(* Logix 5000 project; controller TFF vendor 1 type 14 code 107 rev 34.11; software revision 34.03; part 19 of 36 *)
(* tags used below, declared in another part *)
   AddressPump1 : DINT;   // Temp Address for Pump 1
   AddressPump2 : DINT;   // Temp Address for Pump 2
   Index : DINT;   // Index
   AlarmAnalog : AlarmAnalog[50];   // Analog Alarm Array
   AlarmControl : AlarmControl;   // Alarm Control
   AlarmDeviation : AlarmDeviation[20];   // Control Loop Deviation Alarm Array
   AnalogPoint : AnalogInput[50];   // Analog Input Array
   ControlLoop : ControlLoop[20];   // Control Loop Array
   ControlLoop_FeedBagLevel : ALIAS FOR ControlLoop[2];   // Feed Bag Level Control Loop
   ControlLoop_FeedBagLevelAlarm : ALIAS FOR AlarmDeviation[2];   // Feed Bag Level Control Loop Deviation Alarm
   ControlLoop_FeedPump : ALIAS FOR ControlLoop[1];   // Feed Pump Control Loop
   ControlLoop_FeedPumpAlarm : ALIAS FOR AlarmDeviation[1];   // Feed Pump Control Loop Deviation Alarm
   ControlLoop_PCV001 : ALIAS FOR ControlLoop[3];   // PCV001 Control Loop
   ControlLoop_PCV001Alarm : ALIAS FOR AlarmDeviation[3];   // PCV001 Control Loop Deviation Alarm
   ControlLoop_PCV101 : ALIAS FOR ControlLoop[5];   // PCV101 Control Loop
   ControlLoop_PCV101Alarm : ALIAS FOR AlarmDeviation[5];   // PCV101 Control Loop Deviation Alarm
   Drive : Drive[11];   // Drives Array
   PCV001 : ALIAS FOR AnalogPoint[3];   // Retentate Pressure Control Valve Position
   PCV101 : ALIAS FOR AnalogPoint[4];   // Filtrate Pressure Control Valve Position
   Timers : Timers[22];   // Timer Array
(* Process, continued *)

ROUTINE Alarm_Analog   (* ladder *)
// Analog Alarm Routine
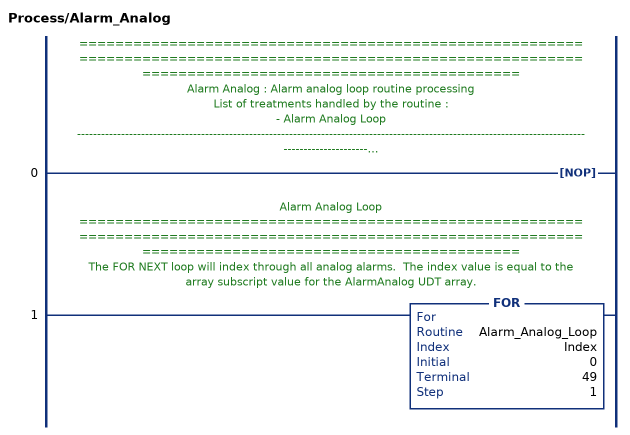
   // ==========================================================================================================================================================
   //                                                                                                                 Alarm Analog : Alarm analog loop routine processing
   //                                                     List of treatments handled by the routine :
   //                                                          - Alarm Analog Loop
   //                                                     -----------------------------------------------------------------------------------------------------------------------------------------------------
   //                                                     History
   //                                                          2019-AUG-13 - Actemium - B. Roch - Initial version for Candidate Release 3.00.00.00.a
   // ==========================================================================================================================================================
   0: NOP();
   // Alarm Analog Loop
   // ==========================================================================================================================================================
   // The FOR NEXT loop will index through all analog alarms.  The index value is equal to the array subscript value for the AlarmAnalog UDT array.
   1: FOR(Alarm_Analog_Loop,Index,0,49,1);
END_ROUTINE

ROUTINE Alarm_Analog_Loop   (* ladder *)
// Analog Alarm Routine
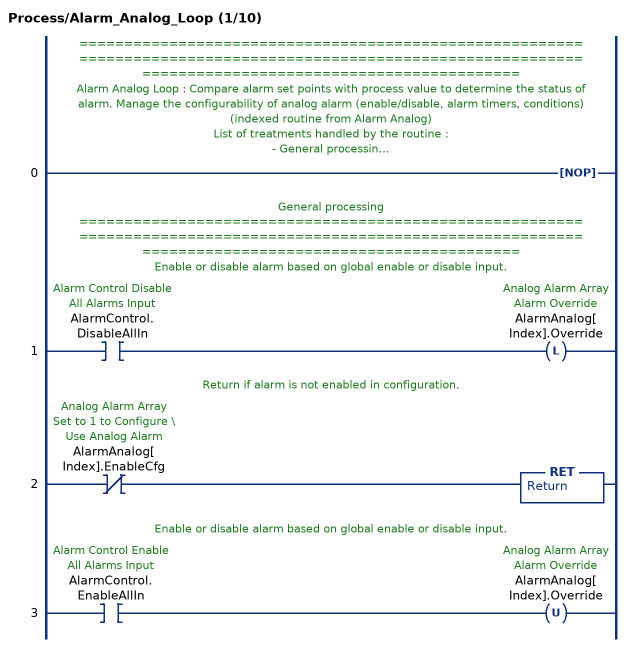
   // ==========================================================================================================================================================
   //           Alarm Analog Loop : Compare alarm set points with process value to determine the status of alarm. Manage the configurability of analog alarm (enable/disable, alarm timers, conditions)
   //                                                                                                                             (indexed routine from Alarm Analog)
   //                                                     List of treatments handled by the routine :
   //                                                          - General processing
   //                                                          - Alarm Acknowledged status
   //                                                          - Alarm conditioned on pump operating status
   //                                                          - Alarm LOLO processing
   //                                                          - Alarm LO processing
   //                                                          - Alarm HI processing
   //                                                          - Alarm HIHI processing
   //                                                          - Alarm status processing
   //                                                     -----------------------------------------------------------------------------------------------------------------------------------------------------
   //                                                     History
   //                                                          2019-AUG-13 - Actemium - B. Roch - Initial version for Candidate Release 3.00.00.00.a
   // ==========================================================================================================================================================
   0: NOP();
   // General processing
   // ==========================================================================================================================================================
   // Enable or disable alarm based on global enable or disable input.
   1: XIC(AlarmControl.DisableAllIn)OTL(AlarmAnalog[Index].Override);
   // Return if alarm is not enabled in configuration.
   2: XIO(AlarmAnalog[Index].EnableCfg)RET();
   // Enable or disable alarm based on global enable or disable input.
   3: XIC(AlarmControl.EnableAllIn)OTU(AlarmAnalog[Index].Override);
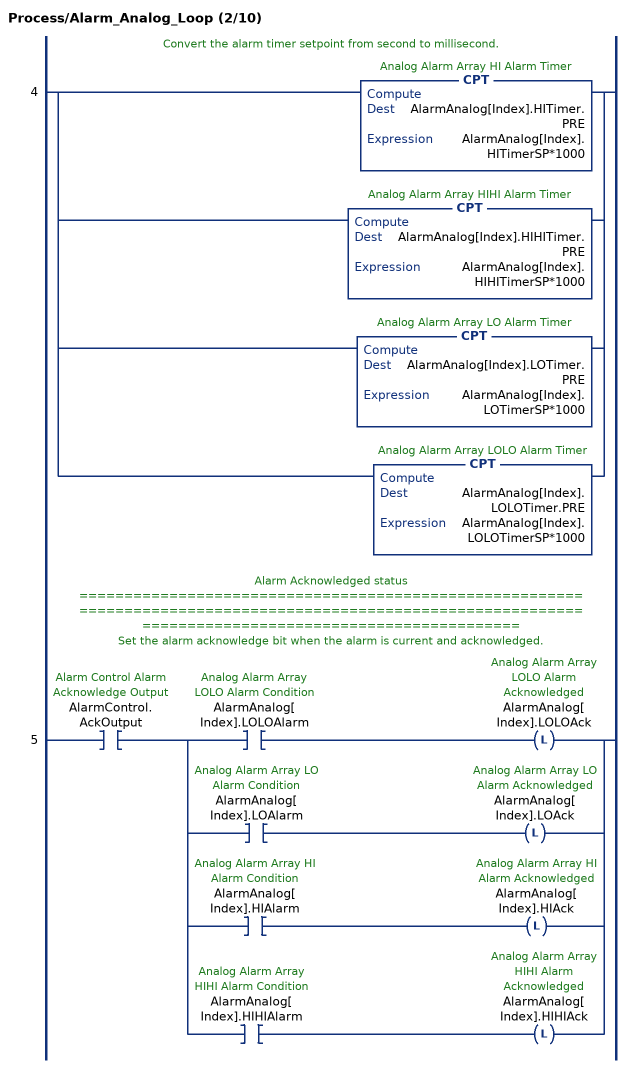
   // Convert the alarm timer setpoint from second to millisecond.
   4: [CPT(AlarmAnalog[Index].HITimer.PRE,AlarmAnalog[Index].HITimerSP*1000) ,CPT(AlarmAnalog[Index].HIHITimer.PRE,AlarmAnalog[Index].HIHITimerSP*1000) ,CPT(AlarmAnalog[Index].LOTimer.PRE,AlarmAnalog[Index].LOTimerSP*1000) ,CPT(AlarmAnalog[Index].LOLOTimer.PRE,AlarmAnalog[Index].LOLOTimerSP*1000) ];
   // Alarm Acknowledged status
   // ==========================================================================================================================================================
   // Set the alarm acknowledge bit when the alarm is current and acknowledged.
   5: XIC(AlarmControl.AckOutput)[XIC(AlarmAnalog[Index].LOLOAlarm) OTL(AlarmAnalog[Index].LOLOAck) ,XIC(AlarmAnalog[Index].LOAlarm) OTL(AlarmAnalog[Index].LOAck) ,XIC(AlarmAnalog[Index].HIAlarm) OTL(AlarmAnalog[Index].HIAck) ,XIC(AlarmAnalog[Index].HIHIAlarm) OTL(AlarmAnalog[Index].HIHIAck) ];
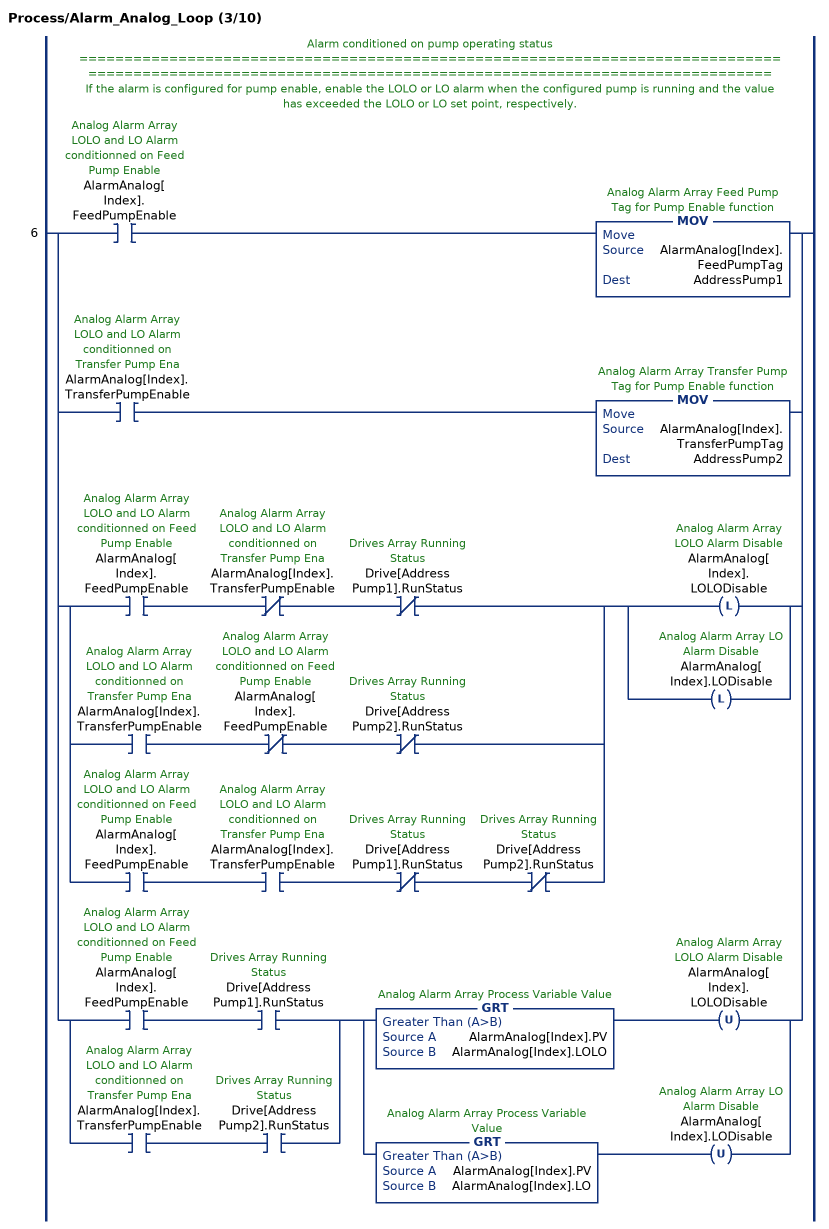
   // Alarm conditioned on pump operating status
   // ==========================================================================================================================================================
   // If the alarm is configured for pump enable, enable the LOLO or LO alarm when the configured pump is running and the value has exceeded the LOLO or LO set point, respectively.
   6: [XIC(AlarmAnalog[Index].FeedPumpEnable) MOV(AlarmAnalog[Index].FeedPumpTag,AddressPump1) ,XIC(AlarmAnalog[Index].TransferPumpEnable) MOV(AlarmAnalog[Index].TransferPumpTag,AddressPump2) ,[XIC(AlarmAnalog[Index].FeedPumpEnable) XIO(AlarmAnalog[Index].TransferPumpEnable) XIO(Drive[AddressPump1].RunStatus) ,XIC(AlarmAnalog[Index].TransferPumpEnable) XIO(AlarmAnalog[Index].FeedPumpEnable) XIO(Drive[AddressPump2].RunStatus) ,XIC(AlarmAnalog[Index].FeedPumpEnable) XIC(AlarmAnalog[Index].TransferPumpEnable) XIO(Drive[AddressPump1].RunStatus) XIO(Drive[AddressPump2].RunStatus) ] [OTL(AlarmAnalog[Index].LOLODisable) ,OTL(AlarmAnalog[Index].LODisable) ] ,[XIC(AlarmAnalog[Index].FeedPumpEnable) XIC(Drive[AddressPump1].RunStatus) ,XIC(AlarmAnalog[Index].TransferPumpEnable) XIC(Drive[AddressPump2].RunStatus) ] [GRT(AlarmAnalog[Index].PV,AlarmAnalog[Index].LOLO) OTU(AlarmAnalog[Index].LOLODisable) ,GRT(AlarmAnalog[Index].PV,AlarmAnalog[Index].LO) OTU(AlarmAnalog[Index].LODisable) ] ];
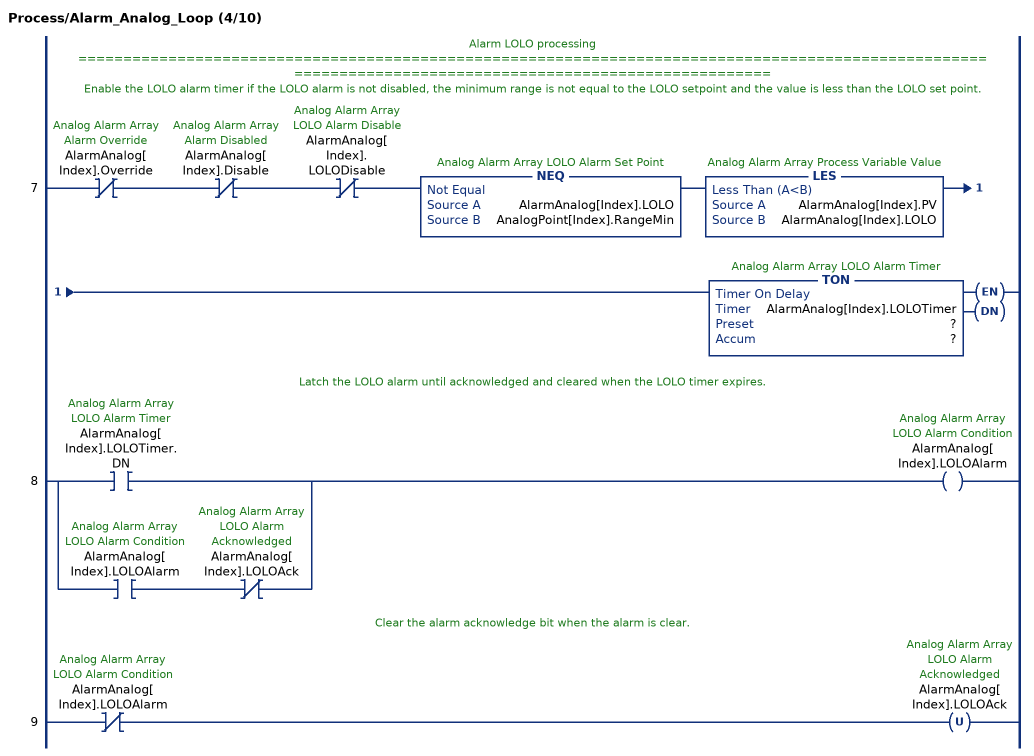
   // Alarm LOLO processing
   // ==========================================================================================================================================================
   // Enable the LOLO alarm timer if the LOLO alarm is not disabled, the minimum range is not equal to the LOLO setpoint and the value is less than the LOLO set point.
   7: XIO(AlarmAnalog[Index].Override)XIO(AlarmAnalog[Index].Disable)XIO(AlarmAnalog[Index].LOLODisable)NEQ(AlarmAnalog[Index].LOLO,AnalogPoint[Index].RangeMin)LES(AlarmAnalog[Index].PV,AlarmAnalog[Index].LOLO)TON(AlarmAnalog[Index].LOLOTimer,?,?);
   // Latch the LOLO alarm until acknowledged and cleared when the LOLO timer expires.
   8: [XIC(AlarmAnalog[Index].LOLOTimer.DN) ,XIC(AlarmAnalog[Index].LOLOAlarm) XIO(AlarmAnalog[Index].LOLOAck) ]OTE(AlarmAnalog[Index].LOLOAlarm);
   // Clear the alarm acknowledge bit when the alarm is clear.
   9: XIO(AlarmAnalog[Index].LOLOAlarm)OTU(AlarmAnalog[Index].LOLOAck);
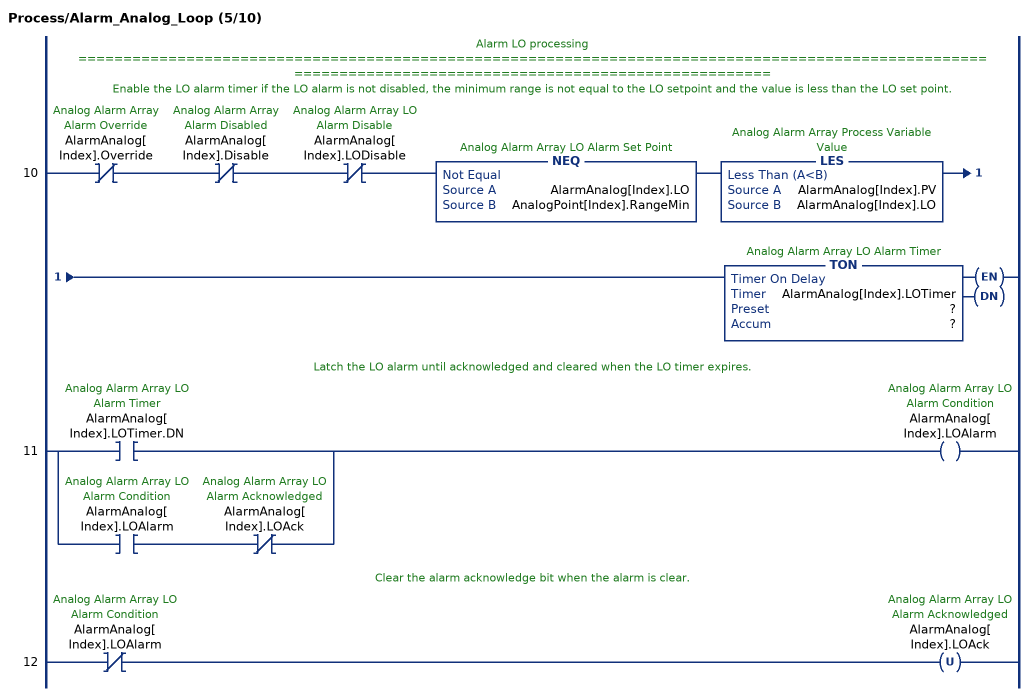
   // Alarm LO processing
   // ==========================================================================================================================================================
   // Enable the LO alarm timer if the LO alarm is not disabled, the minimum range is not equal to the LO setpoint and the value is less than the LO set point.
   10: XIO(AlarmAnalog[Index].Override)XIO(AlarmAnalog[Index].Disable)XIO(AlarmAnalog[Index].LODisable)NEQ(AlarmAnalog[Index].LO,AnalogPoint[Index].RangeMin)LES(AlarmAnalog[Index].PV,AlarmAnalog[Index].LO)TON(AlarmAnalog[Index].LOTimer,?,?);
   // Latch the LO alarm until acknowledged and cleared when the LO timer expires.
   11: [XIC(AlarmAnalog[Index].LOTimer.DN) ,XIC(AlarmAnalog[Index].LOAlarm) XIO(AlarmAnalog[Index].LOAck) ]OTE(AlarmAnalog[Index].LOAlarm);
   // Clear the alarm acknowledge bit when the alarm is clear.
   12: XIO(AlarmAnalog[Index].LOAlarm)OTU(AlarmAnalog[Index].LOAck);
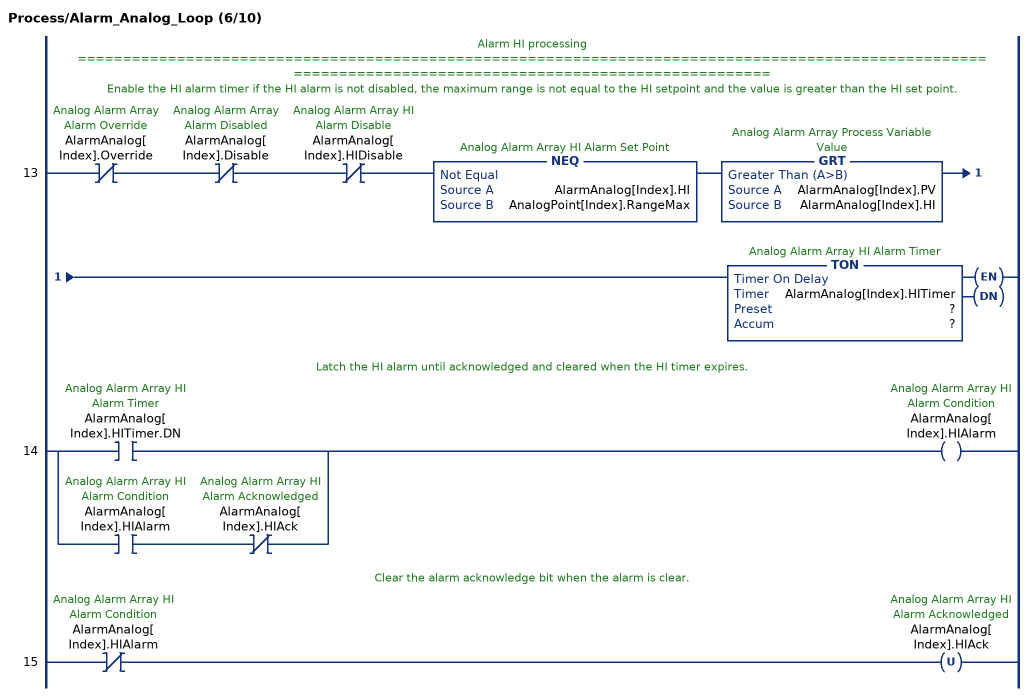
   // Alarm HI processing
   // ==========================================================================================================================================================
   // Enable the HI alarm timer if the HI alarm is not disabled, the maximum range is not equal to the HI setpoint and the value is greater than the HI set point.
   13: XIO(AlarmAnalog[Index].Override)XIO(AlarmAnalog[Index].Disable)XIO(AlarmAnalog[Index].HIDisable)NEQ(AlarmAnalog[Index].HI,AnalogPoint[Index].RangeMax)GRT(AlarmAnalog[Index].PV,AlarmAnalog[Index].HI)TON(AlarmAnalog[Index].HITimer,?,?);
   // Latch the HI alarm until acknowledged and cleared when the HI timer expires.
   14: [XIC(AlarmAnalog[Index].HITimer.DN) ,XIC(AlarmAnalog[Index].HIAlarm) XIO(AlarmAnalog[Index].HIAck) ]OTE(AlarmAnalog[Index].HIAlarm);
   // Clear the alarm acknowledge bit when the alarm is clear.
   15: XIO(AlarmAnalog[Index].HIAlarm)OTU(AlarmAnalog[Index].HIAck);
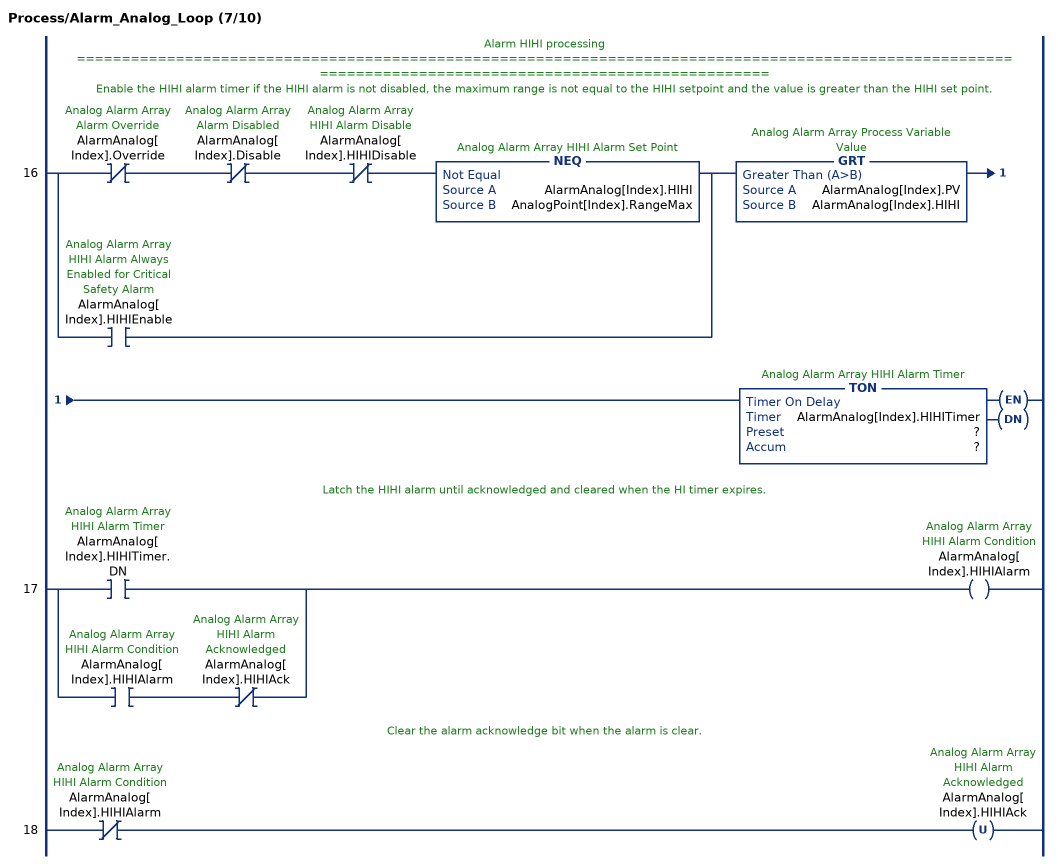
   // Alarm HIHI processing
   // ==========================================================================================================================================================
   // Enable the HIHI alarm timer if the HIHI alarm is not disabled, the maximum range is not equal to the HIHI setpoint and the value is greater than the HIHI set point.
   16: [XIO(AlarmAnalog[Index].Override) XIO(AlarmAnalog[Index].Disable) XIO(AlarmAnalog[Index].HIHIDisable) NEQ(AlarmAnalog[Index].HIHI,AnalogPoint[Index].RangeMax) ,XIC(AlarmAnalog[Index].HIHIEnable) ]GRT(AlarmAnalog[Index].PV,AlarmAnalog[Index].HIHI)TON(AlarmAnalog[Index].HIHITimer,?,?);
   // Latch the HIHI alarm until acknowledged and cleared when the HI timer expires.
   17: [XIC(AlarmAnalog[Index].HIHITimer.DN) ,XIC(AlarmAnalog[Index].HIHIAlarm) XIO(AlarmAnalog[Index].HIHIAck) ]OTE(AlarmAnalog[Index].HIHIAlarm);
   // Clear the alarm acknowledge bit when the alarm is clear.
   18: XIO(AlarmAnalog[Index].HIHIAlarm)OTU(AlarmAnalog[Index].HIHIAck);
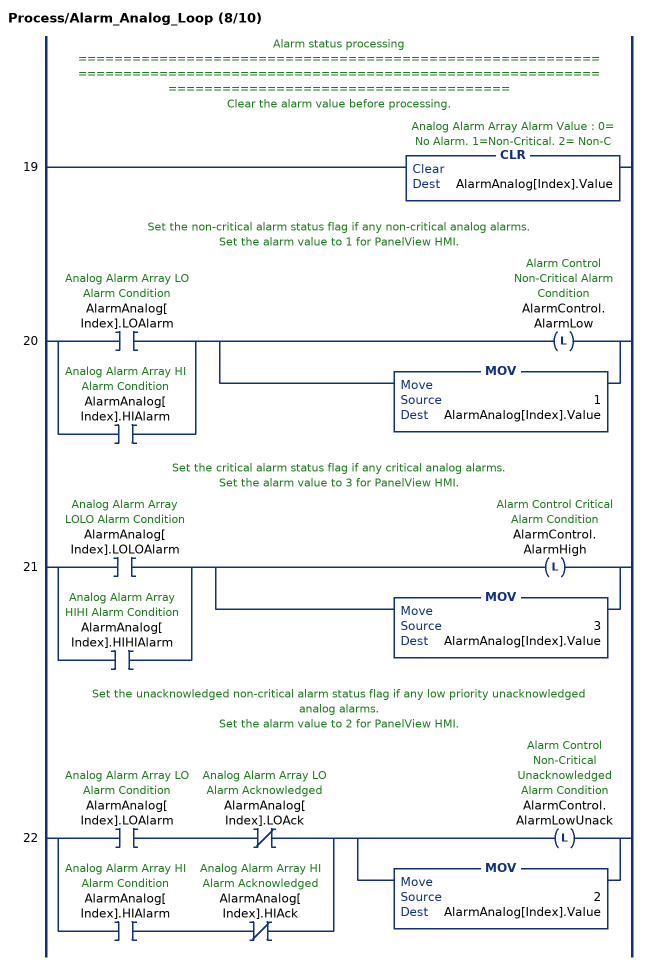
   // Alarm status processing
   // ==========================================================================================================================================================
   // Clear the alarm value before processing.
   19: CLR(AlarmAnalog[Index].Value);
   // Set the non-critical alarm status flag if any non-critical analog alarms.
   // Set the alarm value to 1 for PanelView HMI.
   20: [XIC(AlarmAnalog[Index].LOAlarm) ,XIC(AlarmAnalog[Index].HIAlarm) ][OTL(AlarmControl.AlarmLow) ,MOV(1,AlarmAnalog[Index].Value) ];
   // Set the critical alarm status flag if any critical analog alarms.
   // Set the alarm value to 3 for PanelView HMI.
   21: [XIC(AlarmAnalog[Index].LOLOAlarm) ,XIC(AlarmAnalog[Index].HIHIAlarm) ][OTL(AlarmControl.AlarmHigh) ,MOV(3,AlarmAnalog[Index].Value) ];
   // Set the unacknowledged non-critical alarm status flag if any low priority unacknowledged analog alarms.
   // Set the alarm value to 2 for PanelView HMI.
   22: [XIC(AlarmAnalog[Index].LOAlarm) XIO(AlarmAnalog[Index].LOAck) ,XIC(AlarmAnalog[Index].HIAlarm) XIO(AlarmAnalog[Index].HIAck) ][OTL(AlarmControl.AlarmLowUnack) ,MOV(2,AlarmAnalog[Index].Value) ];
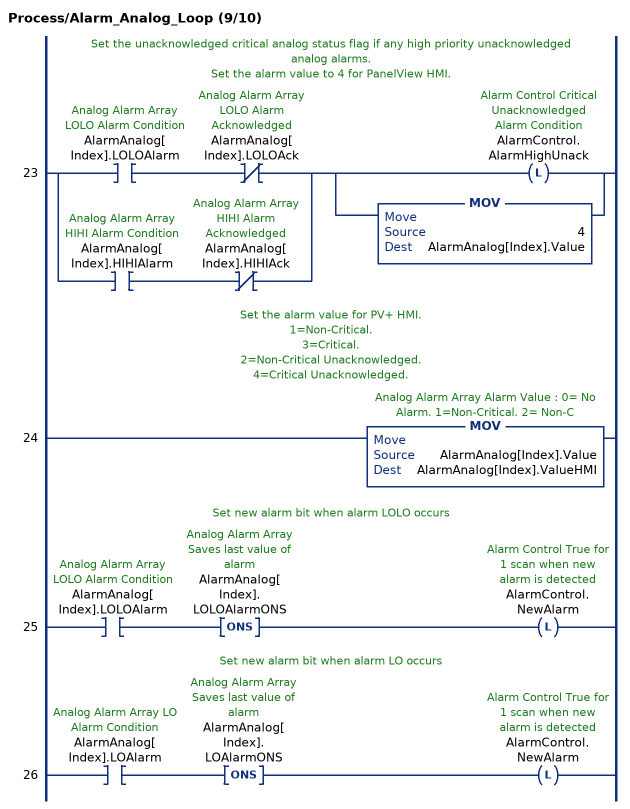
   // Set the unacknowledged critical analog status flag if any high priority unacknowledged analog alarms.
   // Set the alarm value to 4 for PanelView HMI.
   23: [XIC(AlarmAnalog[Index].LOLOAlarm) XIO(AlarmAnalog[Index].LOLOAck) ,XIC(AlarmAnalog[Index].HIHIAlarm) XIO(AlarmAnalog[Index].HIHIAck) ][OTL(AlarmControl.AlarmHighUnack) ,MOV(4,AlarmAnalog[Index].Value) ];
   // Set the alarm value for PV+ HMI.
   // 1=Non-Critical.
   // 3=Critical.
   // 2=Non-Critical Unacknowledged.
   // 4=Critical Unacknowledged.
   24: MOV(AlarmAnalog[Index].Value,AlarmAnalog[Index].ValueHMI);
   // Set new alarm bit when alarm LOLO occurs
   25: XIC(AlarmAnalog[Index].LOLOAlarm)ONS(AlarmAnalog[Index].LOLOAlarmONS)OTL(AlarmControl.NewAlarm);
   // Set new alarm bit when alarm LO occurs
   26: XIC(AlarmAnalog[Index].LOAlarm)ONS(AlarmAnalog[Index].LOAlarmONS)OTL(AlarmControl.NewAlarm);
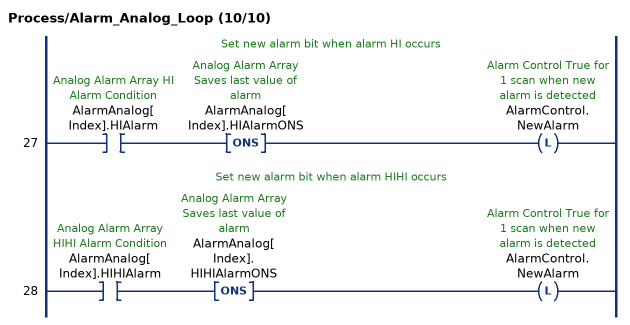
   // Set new alarm bit when alarm HI occurs
   27: XIC(AlarmAnalog[Index].HIAlarm)ONS(AlarmAnalog[Index].HIAlarmONS)OTL(AlarmControl.NewAlarm);
   // Set new alarm bit when alarm HIHI occurs
   28: XIC(AlarmAnalog[Index].HIHIAlarm)ONS(AlarmAnalog[Index].HIHIAlarmONS)OTL(AlarmControl.NewAlarm);
END_ROUTINE

ROUTINE Alarm_Deviation   (* ladder *)
// Deviation Alarm Routine
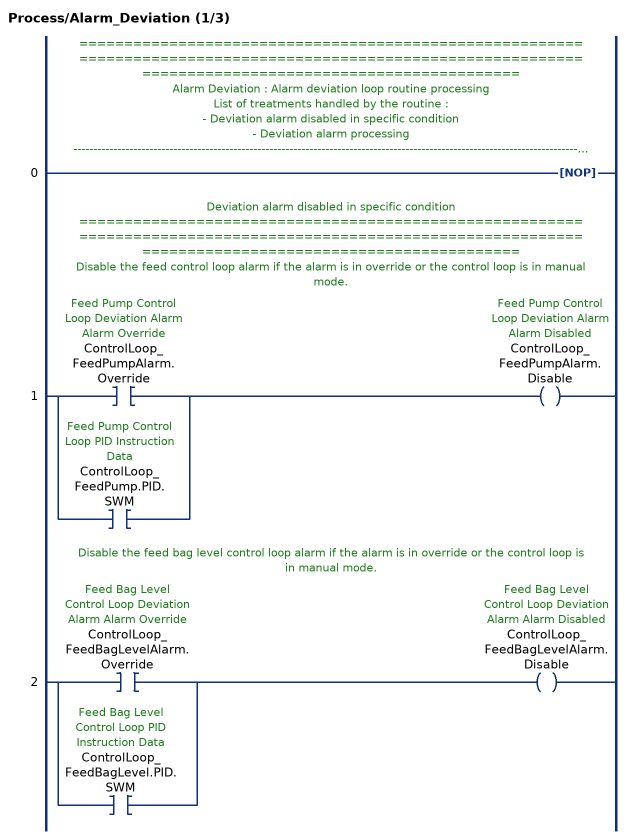
   // ==========================================================================================================================================================
   //                                                                                                         Alarm Deviation : Alarm deviation loop routine processing
   //                                                     List of treatments handled by the routine :
   //                                                          - Deviation alarm disabled in specific condition
   //                                                          - Deviation alarm processing
   //                                                     -----------------------------------------------------------------------------------------------------------------------------------------------------
   //                                                     History
   //                                                          2019-AUG-13 - Actemium - B. Roch - Initial version for Candidate Release 3.00.00.00.a
   //                                                          2019-SEP-26 - Actemium - B. Roch - Modification for Candidate Release 3.00.00.00.c
   //                                 - Change activation condition for PCV alarm deviation
   // ==========================================================================================================================================================
   0: NOP();
   // Deviation alarm disabled in specific condition
   // ==========================================================================================================================================================
   // Disable the feed control loop alarm if the alarm is in override or the control loop is in manual mode.
   1: [XIC(ControlLoop_FeedPumpAlarm.Override) ,XIC(ControlLoop_FeedPump.PID.SWM) ]OTE(ControlLoop_FeedPumpAlarm.Disable);
   // Disable the feed bag level control loop alarm if the alarm is in override or the control loop is in manual mode.
   2: [XIC(ControlLoop_FeedBagLevelAlarm.Override) ,XIC(ControlLoop_FeedBagLevel.PID.SWM) ]OTE(ControlLoop_FeedBagLevelAlarm.Disable);
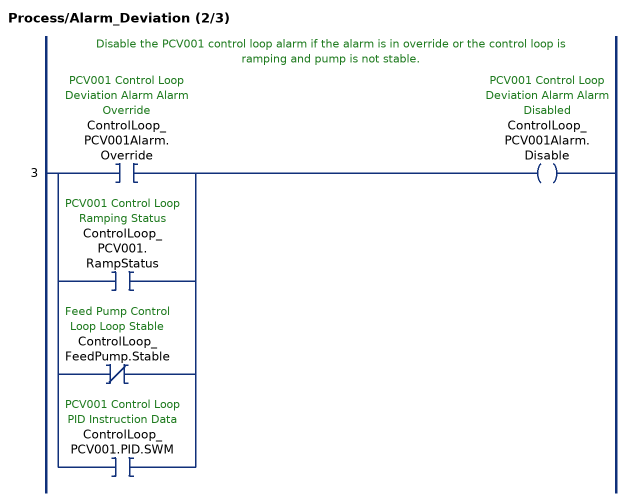
   // Disable the PCV001 control loop alarm if the alarm is in override or the control loop is ramping and pump is not stable.
   3: [XIC(ControlLoop_PCV001Alarm.Override) ,XIC(ControlLoop_PCV001.RampStatus) ,XIO(ControlLoop_FeedPump.Stable) ,XIC(ControlLoop_PCV001.PID.SWM) ]OTE(ControlLoop_PCV001Alarm.Disable);
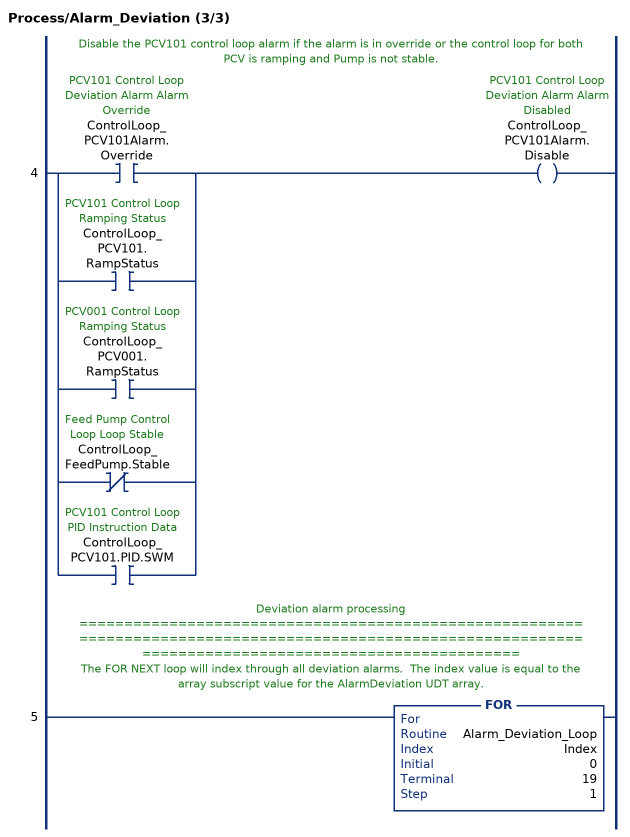
   // Disable the PCV101 control loop alarm if the alarm is in override or the control loop for both PCV is ramping and Pump is not stable.
   4: [XIC(ControlLoop_PCV101Alarm.Override) ,XIC(ControlLoop_PCV101.RampStatus) ,XIC(ControlLoop_PCV001.RampStatus) ,XIO(ControlLoop_FeedPump.Stable) ,XIC(ControlLoop_PCV101.PID.SWM) ]OTE(ControlLoop_PCV101Alarm.Disable);
   // Deviation alarm processing
   // ==========================================================================================================================================================
   // The FOR NEXT loop will index through all deviation alarms.  The index value is equal to the array subscript value for the AlarmDeviation UDT array.
   5: FOR(Alarm_Deviation_Loop,Index,0,19,1);
END_ROUTINE

ROUTINE Alarm_Deviation_Loop   (* ladder *)
// Deviation Alarm Routine
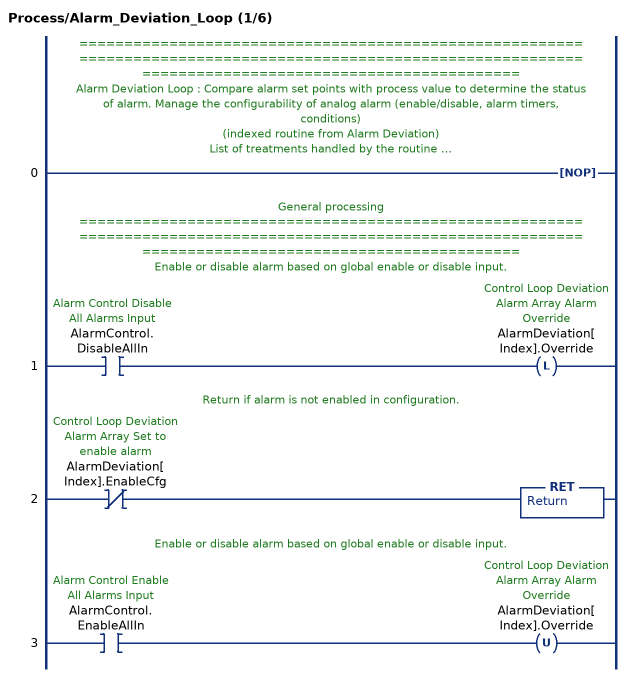
   // ==========================================================================================================================================================
   //        Alarm Deviation Loop : Compare alarm set points with process value to determine the status of alarm. Manage the configurability of analog alarm (enable/disable, alarm timers, conditions)
   //                                                                                                                             (indexed routine from Alarm Deviation)
   //                                                     List of treatments handled by the routine :
   //                                                          - General processing
   //                                                          - Alarm Acknowledged status
   //                                                          - Alarm HI processing
   //                                                          - Alarm HIHI processing
   //                                                          - Alarm status processing
   //                                                     -----------------------------------------------------------------------------------------------------------------------------------------------------
   //                                                     History
   //                                                          2019-AUG-13 - Actemium - B. Roch - Initial version for Candidate Release 3.00.00.00.a
   // ==========================================================================================================================================================
   0: NOP();
   // General processing
   // ==========================================================================================================================================================
   // Enable or disable alarm based on global enable or disable input.
   1: XIC(AlarmControl.DisableAllIn)OTL(AlarmDeviation[Index].Override);
   // Return if alarm is not enabled in configuration.
   2: XIO(AlarmDeviation[Index].EnableCfg)RET();
   // Enable or disable alarm based on global enable or disable input.
   3: XIC(AlarmControl.EnableAllIn)OTU(AlarmDeviation[Index].Override);
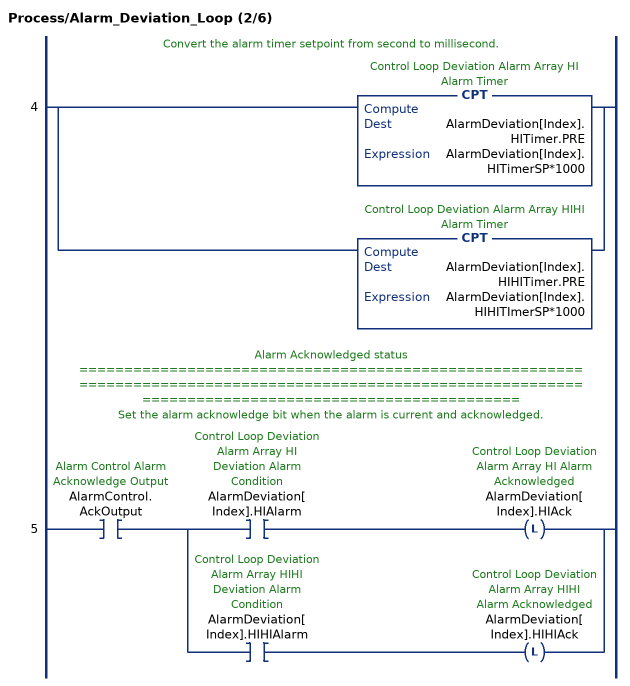
   // Convert the alarm timer setpoint from second to millisecond.
   4: [CPT(AlarmDeviation[Index].HITimer.PRE,AlarmDeviation[Index].HITimerSP*1000) ,CPT(AlarmDeviation[Index].HIHITimer.PRE,AlarmDeviation[Index].HIHITImerSP*1000) ];
   // Alarm Acknowledged status
   // ==========================================================================================================================================================
   // Set the alarm acknowledge bit when the alarm is current and acknowledged.
   5: XIC(AlarmControl.AckOutput)[XIC(AlarmDeviation[Index].HIAlarm) OTL(AlarmDeviation[Index].HIAck) ,XIC(AlarmDeviation[Index].HIHIAlarm) OTL(AlarmDeviation[Index].HIHIAck) ];
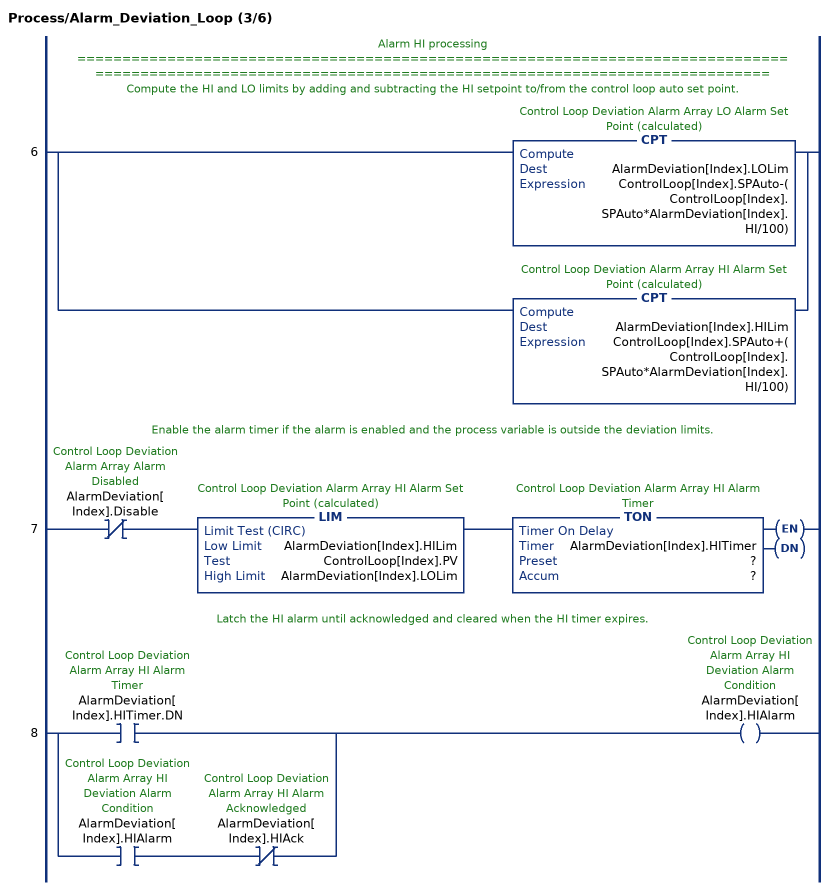
   // Alarm HI processing
   // ==========================================================================================================================================================
   // Compute the HI and LO limits by adding and subtracting the HI setpoint to/from the control loop auto set point.
   6: [CPT(AlarmDeviation[Index].LOLim,ControlLoop[Index].SPAuto-(ControlLoop[Index].SPAuto*AlarmDeviation[Index].HI/100)) ,CPT(AlarmDeviation[Index].HILim,ControlLoop[Index].SPAuto+(ControlLoop[Index].SPAuto*AlarmDeviation[Index].HI/100)) ];
   // Enable the alarm timer if the alarm is enabled and the process variable is outside the deviation limits.
   7: XIO(AlarmDeviation[Index].Disable)LIM(AlarmDeviation[Index].HILim,ControlLoop[Index].PV,AlarmDeviation[Index].LOLim)TON(AlarmDeviation[Index].HITimer,?,?);
   // Latch the HI alarm until acknowledged and cleared when the HI timer expires.
   8: [XIC(AlarmDeviation[Index].HITimer.DN) ,XIC(AlarmDeviation[Index].HIAlarm) XIO(AlarmDeviation[Index].HIAck) ]OTE(AlarmDeviation[Index].HIAlarm);
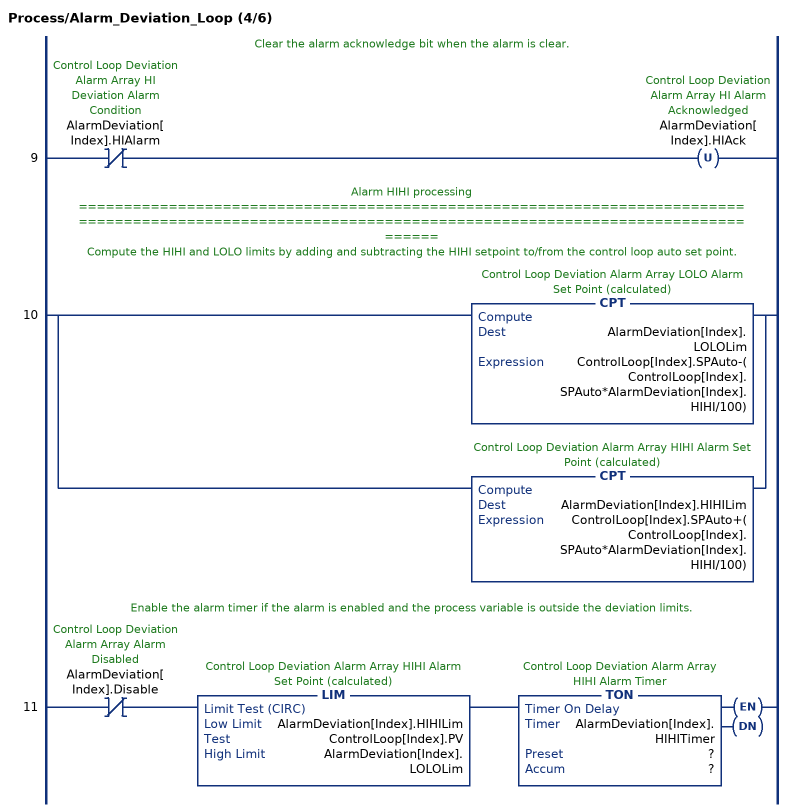
   // Clear the alarm acknowledge bit when the alarm is clear.
   9: XIO(AlarmDeviation[Index].HIAlarm)OTU(AlarmDeviation[Index].HIAck);
   // Alarm HIHI processing
   // ==========================================================================================================================================================
   // Compute the HIHI and LOLO limits by adding and subtracting the HIHI setpoint to/from the control loop auto set point.
   10: [CPT(AlarmDeviation[Index].LOLOLim,ControlLoop[Index].SPAuto-(ControlLoop[Index].SPAuto*AlarmDeviation[Index].HIHI/100)) ,CPT(AlarmDeviation[Index].HIHILim,ControlLoop[Index].SPAuto+(ControlLoop[Index].SPAuto*AlarmDeviation[Index].HIHI/100)) ];
   // Enable the alarm timer if the alarm is enabled and the process variable is outside the deviation limits.
   11: XIO(AlarmDeviation[Index].Disable)LIM(AlarmDeviation[Index].HIHILim,ControlLoop[Index].PV,AlarmDeviation[Index].LOLOLim)TON(AlarmDeviation[Index].HIHITimer,?,?);
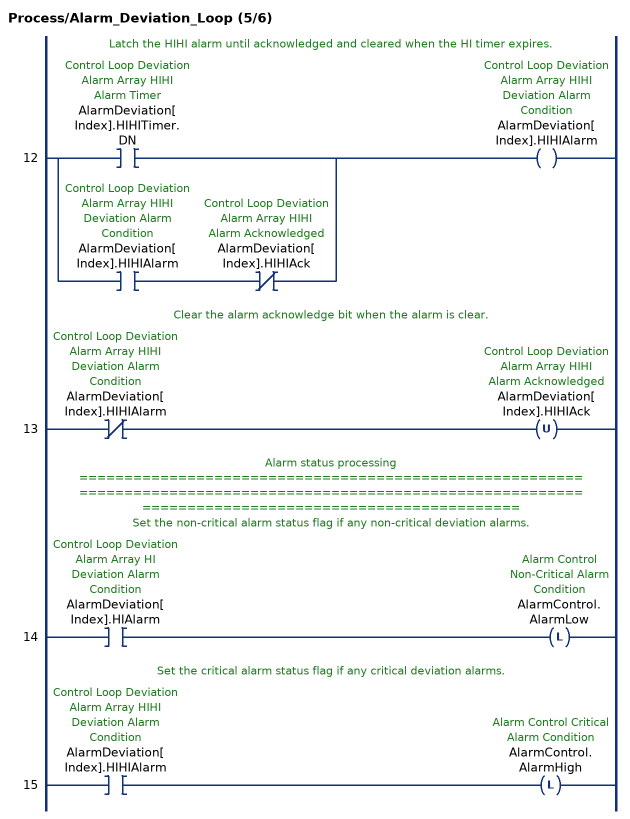
   // Latch the HIHI alarm until acknowledged and cleared when the HI timer expires.
   12: [XIC(AlarmDeviation[Index].HIHITimer.DN) ,XIC(AlarmDeviation[Index].HIHIAlarm) XIO(AlarmDeviation[Index].HIHIAck) ]OTE(AlarmDeviation[Index].HIHIAlarm);
   // Clear the alarm acknowledge bit when the alarm is clear.
   13: XIO(AlarmDeviation[Index].HIHIAlarm)OTU(AlarmDeviation[Index].HIHIAck);
   // Alarm status processing
   // ==========================================================================================================================================================
   // Set the non-critical alarm status flag if any non-critical deviation alarms.
   14: XIC(AlarmDeviation[Index].HIAlarm)OTL(AlarmControl.AlarmLow);
   // Set the critical alarm status flag if any critical deviation alarms.
   15: XIC(AlarmDeviation[Index].HIHIAlarm)OTL(AlarmControl.AlarmHigh);
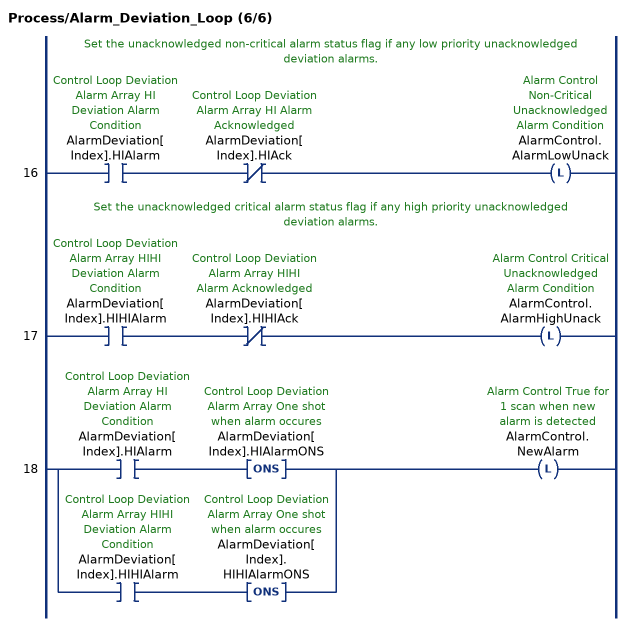
   // Set the unacknowledged non-critical alarm status flag if any low priority unacknowledged deviation alarms.
   16: XIC(AlarmDeviation[Index].HIAlarm)XIO(AlarmDeviation[Index].HIAck)OTL(AlarmControl.AlarmLowUnack);
   // Set the unacknowledged critical alarm status flag if any high priority unacknowledged deviation alarms.
   17: XIC(AlarmDeviation[Index].HIHIAlarm)XIO(AlarmDeviation[Index].HIHIAck)OTL(AlarmControl.AlarmHighUnack);
   18: [XIC(AlarmDeviation[Index].HIAlarm) ONS(AlarmDeviation[Index].HIAlarmONS) ,XIC(AlarmDeviation[Index].HIHIAlarm) ONS(AlarmDeviation[Index].HIHIAlarmONS) ]OTL(AlarmControl.NewAlarm);
END_ROUTINE
